// TIA Portal V20 export
// export: Created 2026-10-20T12:46:59.9047324Z, ExportSetting WithDefaults, DisplayName Totally Integrated Automation Portal, DisplayVersion V20 Update 6, DisplayName TIA Portal Openness, DisplayVersion V20 Update 6, DisplayName TIA Portal Version Control Interface, DisplayVersion V20 Update 6, DisplayName SINAMICS Startdrive Advanced, DisplayVersion V20 SP1, DisplayName SINAMICS Startdrive G130, G150, S120, S150, SINAMICS MV, G220, S200, S210, DisplayVersion V20 SP1, DisplayName SINAMICS Startdrive G110M, G120, G120C, G120D, G120P, G115D, DisplayVersion V20 SP1, DisplayName STEP 7 Professional, DisplayVersion V20 Update 6, DisplayName STEP 7 Safety, DisplayVersion V20 Update 2, DisplayName WinCC Basic/Comfort/Advanced, DisplayVersion V20 Update 6, DisplayName WinCC Unified, DisplayVersion V20 Update 6
FUNCTION "FindIntField" : Int   // FC18, SCL
{ S7_Optimized_Access := 'TRUE' }
VERSION : 0.1
// stored: AutoNumber true, IsIECCheckEnabled false, SetENOAutomatically false, UDAEnableTagReadback false
   VAR_INPUT
      FieldName : String;
      JsonStr : String;
   END_VAR
   VAR_TEMP
      searchStr : String;
      foundPos : Int;
      valueStr : String;
      delimPos : Int;
   END_VAR
BEGIN
   // Set up the search pattern, e.g. '"id":'
   #searchStr := CONCAT(IN1 := '"', IN2 := #FieldName);
   #searchStr := CONCAT(IN1 := #searchStr, IN2 := '" :');

   // Search the field
   #foundPos := FIND(IN1 := #JsonStr, IN2 := #searchStr);

   IF #foundPos > 0 THEN
       // Try to find a comma after the value
       #delimPos := FIND(
                         IN1 := MID(IN := #JsonStr, P := #foundPos + LEN(#searchStr), L := 10),
                         IN2 := ','
       );

       // If there is no comma, try to find the closing brace '}'
       IF #delimPos = 0 THEN
           #delimPos := FIND(
                             IN1 := MID(IN := #JsonStr, P := #foundPos + LEN(#searchStr), L := 10),
                             IN2 := '}'
           );
       END_IF;

       // If you find the end of value, extract the value
       IF #delimPos > 0 THEN
           #valueStr := MID(
                            IN := #JsonStr,
                            P := #foundPos + LEN(#searchStr),
                            L := #delimPos - 1
           );
           #FindIntField := STRING_TO_INT(#valueStr);
           RETURN;
       END_IF;
   END_IF;

   // Default return if not found or error
   #FindIntField := -9999;
END_FUNCTION
